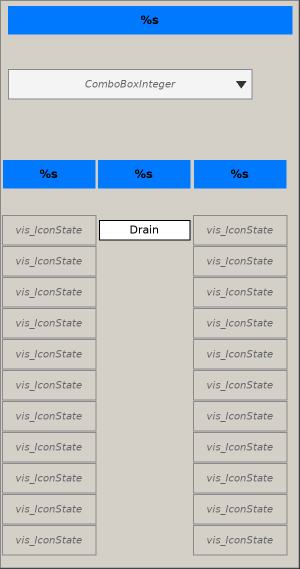
VISUALIZATION vis_FB_ProductionTank  // 300x569
VAR_IN_OUT
	fb: FB_ProductionTank;
END_VAR
    Rectangle (0,0 300x569)
    Textfield (7,5 286x30), "%s", text variable: fb.refElement.sElementID
    RoundedRectangle (99,220 91x20), "Drain"
        OnMouseClick: execute { fb.eReq:=E_Request_List.eDrain; }
    ComboBoxInteger (8,69 244x30), variable: fb.refElement.eState_Long, input disabled if: fb.refElement.bStateUpdate_Limited, text list: 'TextList_StateLong'
    Textfield (97,159 94x30), "%s", text variable: fb.eReq
    Textfield (193,159 94x30), "%s", text variable: fb.eProcess
    Textfield (2,159 94x30), "%s", text variable: fb.refElement.eState_Long, text list: 'TextList_StateLong', text index: fb.refElement.eState_Long
    Frame (2,215 94x30)
        shows vis_IconState(value := fb.refElement.eState_Long, reqValue := E_Element_State_Long.eStandby, text := 'Standby')
    Frame (2,246 94x30)
        shows vis_IconState(value := fb.refElement.eState_Long, reqValue := E_Element_State_Long.eNotClean, text := 'Not Clean')
    Frame (2,277 94x30)
        shows vis_IconState(value := fb.refElement.eState_Long, reqValue := E_Element_State_Long.eCIP_1_Rinzed, text := 'CIP1 Rinzed')
    Frame (2,308 94x30)
        shows vis_IconState(value := fb.refElement.eState_Long, reqValue := E_Element_State_Long.eCIP_2_Deterged, text := 'CIP2 Deterged')
    Frame (2,339 94x30)
        shows vis_IconState(value := fb.refElement.eState_Long, reqValue := E_Element_State_Long.eCIP_3_Deterged_Clean, text := 'CIP3 Deterged +')
    Frame (2,370 94x30)
        shows vis_IconState(value := fb.refElement.eState_Long, reqValue := E_Element_State_Long.eCIP_4_Sanitized, text := 'DisInfected')
    Frame (2,401 94x30)
        shows vis_IconState(value := fb.refElement.eState_Long, reqValue := E_Element_State_Long.eCIP_5_Done, text := 'CIP5 Done')
    Frame (2,432 94x30)
        shows vis_IconState(value := fb.refElement.eState_Long, reqValue := E_Element_State_Long.eWaterReady, text := 'WaterReady')
    Frame (2,463 94x30)
        shows vis_IconState(value := fb.refElement.eState_Long, reqValue := E_Element_State_Long.eReady, text := 'Ready')
    Frame (2,494 94x30)
        shows vis_IconState(value := fb.refElement.eState_Long, reqValue := E_Element_State_Long.eProduction, text := 'Production')
    Frame (2,525 94x30)
        shows vis_IconState(value := fb.refElement.eState_Long, reqValue := E_Element_State_Long.eExpired, text := 'Expired')
    Frame (193,215 94x30)
        shows vis_IconState(value := fb.eProcess, reqValue := E_Element_Process.eDrain, text := 'Draining')
    Frame (193,246 94x30)
        shows vis_IconState(value := fb.eProcess, reqValue := E_Element_Process.eWash_Recycle, text := 'Wash Recycle')
    Frame (193,277 94x30)
        shows vis_IconState(value := fb.eProcess, reqValue := E_Element_Process.eWash_Detergent, text := 'Wash Detergent')
    Frame (193,308 94x30)
        shows vis_IconState(value := fb.eProcess, reqValue := E_Element_Process.eWash_Water_1, text := 'Water 1')
    Frame (193,339 94x30)
        shows vis_IconState(value := fb.eProcess, reqValue := E_Element_Process.eWash_Sani, text := 'Wash DisInfection')
    Frame (193,370 94x30)
        shows vis_IconState(value := fb.eProcess, reqValue := E_Element_Process.eWash_Water_2, text := 'Water')
    Frame (193,401 94x30)
        shows vis_IconState(value := fb.eProcess, reqValue := E_Element_Process.eFill_Water, text := 'Filling Water')
    Frame (193,432 94x30)
        shows vis_IconState(value := fb.eProcess, reqValue := E_Element_Process.eDissolving, text := 'Dissolving')
    Frame (193,463 94x30)
        shows vis_IconState(value := fb.eProcess, reqValue := E_Element_Process.eConnectionToLine, text := 'Conn To Line')
    Frame (193,494 94x30)
        shows vis_IconState(value := fb.eProcess, reqValue := E_Element_Process.eDisconnection, text := 'Wash Detergent')
    Frame (193,525 94x30)
        shows vis_IconState(value := fb.eProcess, reqValue := E_Element_Process.eDrain, text := ' ')
END_VISUALIZATION

(* stored: Version 1.1.0.1, ProductVersion 3.1.4024.15
   Visu vis_FB_ProductionTank: Id {1a282a5f-038c-4014-a3e8-318e8aa55f48} *)
